// TIA Portal V21 export
FUNCTION "FC_ClampPctLad" : Int   // FC111, LAD
TITLE = Ограничение значения пределами (LAD)
{ S7_Optimized_Access := 'TRUE' }
AUTHOR : WTP2
FAMILY : Utils
VERSION : 0.1
// Результат: iIn, ограниченный снизу iMin и сверху iMax (сначала верхний предел, затем нижний). ENO не пишется: ENO = EN.
// stored: AutoNumber false, SetENOAutomatically false
   VAR_INPUT
      iIn : Int;   // Значение
      iMin : Int;   // Нижний предел
      iMax : Int;   // Верхний предел
   END_VAR
BEGIN

REGION Network 1: Значение по умолчанию
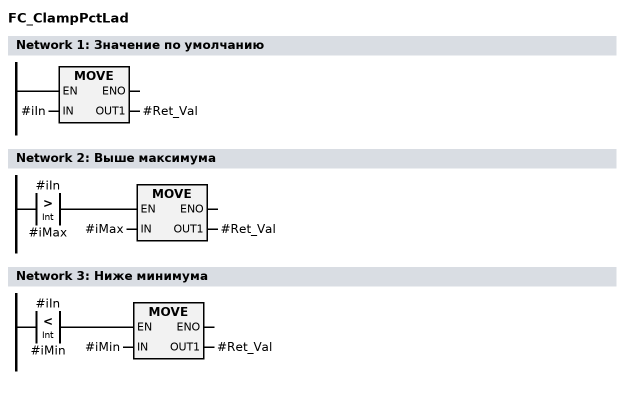
   RUNG wire#powerrail
      Move(in := #iIn, out1 => #Ret_Val)
   END_RUNG
   // the same network as SCL:
   #Ret_Val := #iIn;
END_REGION

REGION Network 2: Выше максимума
   RUNG wire#powerrail
      { S7_Templates := "SrcType := Int" } GT_Contact(in1 := #iIn, in2 := #iMax)
      Move(in := #iMax, out1 => #Ret_Val)
   END_RUNG
   // the same network as SCL:
   IF #iIn > #iMax THEN #Ret_Val := #iMax; END_IF;
END_REGION

REGION Network 3: Ниже минимума
   RUNG wire#powerrail
      { S7_Templates := "SrcType := Int" } LT_Contact(in1 := #iIn, in2 := #iMin)
      Move(in := #iMin, out1 => #Ret_Val)
   END_RUNG
   // the same network as SCL:
   IF #iIn < #iMin THEN #Ret_Val := #iMin; END_IF;
END_REGION
END_FUNCTION
